// TIA Portal V21 export
// export: Created 2026-11-07T15:25:01.9563364Z, ExportSetting WithDefaults, DisplayName Totally Integrated Automation Portal, DisplayVersion V21, DisplayName STEP 7 Professional, DisplayVersion V21, DisplayName STEP 7 Safety, DisplayVersion V21, DisplayName Tech WebApplication, DisplayVersion V21, DisplayName WinCC Basic/Comfort/Advanced, DisplayVersion V21, DisplayName WinCC Unified, DisplayVersion V21
TextList "TL_State"  ListRange=Decimal
  TextListEntry   EntryType=SingleValue, Text="OFF"
  TextListEntry   EntryType=SingleValue, From=1, To=1, Text="INIT"
